(* IEC 61131-3 sources: plcassist-cli/packages/volt-lsp-iec/test-corpus/bakon-nano/Device/Plc Logic/Application/Library Manager/CAA TickUtil, 8 files *)

(* ---- VERSIONCONSTANTS.gvl ---- *)
VAR_GLOBAL
	GC_BYVERSION : BYTE := 1;
	GC_VERSION_1 : BYTE := 0;
END_VAR

(* ---- CONVERTNSECTOTICK.fun ---- *)
FUNCTION CONVERTNSECTOTICK : CAA.TICK
VAR_INPUT
	UDINSECONDS : UDINT;
END_VAR
END_FUNCTION

(* ---- CONVERTTICKTONSEC.fun ---- *)
FUNCTION CONVERTTICKTONSEC : UDINT
VAR_INPUT
	TKTICK : CAA.TICK;
END_VAR
END_FUNCTION

(* ---- CONVERTTICKTOUSEC.fun ---- *)
FUNCTION CONVERTTICKTOUSEC : UDINT
VAR_INPUT
	TKTICK : CAA.TICK;
END_VAR
END_FUNCTION

(* ---- CONVERTUSECTOTICK.fun ---- *)
FUNCTION CONVERTUSECTOTICK : CAA.TICK
VAR_INPUT
	UDIUSECONDS : UDINT;
END_VAR
END_FUNCTION

(* ---- GETELAPSEDTIMEINNSEC.fun ---- *)
FUNCTION GETELAPSEDTIMEINNSEC : UDINT
VAR_INPUT
	TKSTART : CAA.TICK;
END_VAR
END_FUNCTION

(* ---- GETELAPSEDTIMEINUSEC.fun ---- *)
FUNCTION GETELAPSEDTIMEINUSEC : UDINT
VAR_INPUT
	TKSTART : CAA.TICK;
END_VAR
END_FUNCTION

(* ---- GETSUPPLIERVERSION.fun ---- *)
FUNCTION GETSUPPLIERVERSION : WORD
VAR_INPUT
	XDUMMY : BOOL;
END_VAR
END_FUNCTION
